Fanuc KAREL source: ko00082.KL

-- PROVISIONAL review KL for V770-1; original PC SHA256 97795c489b74edf4d54bbb0fc4c0705b0bf3fa318ad31b6fdb71413d2604f282
-- Incomplete behavior may be omitted. Consult companion uncertainty JSON. Do not deploy.
PROGRAM KO00082
%NOLOCKGROUP
BEGIN
  -- UNRESOLVED_PC offsets 5-12; opcodes 9D,23
  -- UNRESOLVED_PC offsets 17-66; opcodes 27,27,49,7E,AD,22,1C,22,31,7E,4A
  -- UNRESOLVED_PC offsets 71-75; opcodes 7F
END KO00082
